Staubli VAL3: renameFrame.pgx

program renameFrame(num x_nIndex)
  local string l_sName
  local bool l_bResult
begin
  l_bResult=userPagePrompt("请输入新的名称：",l_sName)
  if l_bResult
    savedata:fFrameItem[x_nIndex].sName=l_sName
    savedata:libSave()
    delay(0.1)
  endIf
end
